(* IEC 61131-3 sources: kns-pump-station/tests/POUs/Station/FB_ControlSelector_Test, 6 files *)

(* ---- ChangedPulsesOnce.method.decl.st ---- *)
// xChanged — один вызов на смену управления (вход без рывка); без смены — FALSE
METHOD PRIVATE ChangedPulsesOnce
VAR
    fbDut : FB_ControlSelector;          // ФБ под тестом
END_VAR

(* ---- GarbageMethodIsStepped.method.decl.st ---- *)
// Способ вне перечисления — как «Ступенчатое» (E_ControlMethod: безопасный вариант)
METHOD PRIVATE GarbageMethodIsStepped
VAR
    fbDut : FB_ControlSelector;          // ФБ под тестом
    pRaw : POINTER TO INT;             // способ вне перечисления
    eBad  : E_ControlMethod;            // мусор
END_VAR

(* ---- ManualModeAlwaysManual.method.decl.st ---- *)
// 04 §4: в «Ручном» — Manual при любых условиях (защиты действуют блокировками, без запросов); режим вне
// перечисления — как «Ручной»
METHOD PRIVATE ManualModeAlwaysManual
VAR
    fbDut : FB_ControlSelector;          // ФБ под тестом
    pRaw : POINTER TO INT;             // режим вне перечисления
    eBad  : E_StationMode;              // мусор
END_VAR

(* ---- PidNotReadyFallsBackToStepped.method.decl.st ---- *)
// 04 §7.4, PMI-28: выбран ПИД, ПИД не готов — Stepped и условие KNS1.STEP; готов — LevelPid без условия
METHOD PRIVATE PidNotReadyFallsBackToStepped
VAR
    fbDut : FB_ControlSelector;          // ФБ под тестом
END_VAR

(* ---- PrecedenceTable.method.decl.st ---- *)
// 04 §4: старшинство в «Автомате» PowerLost > Restart > DryRunStop > Float > Emergency > LevelPid > Stepped — для
// каждой пары условий побеждает старшее (все 2^5 сочетаний пяти условий при выбранном и готовом ПИД)
METHOD PRIVATE PrecedenceTable
VAR
    fbDut : FB_ControlSelector;          // ФБ под тестом

    uiMask   : UINT;                    // сочетание условий: бит 0 PowerLost … бит 4 Emergency
    eExpect  : E_ControlAct;            // ожидаемое управление
    xAllOk   : BOOL := TRUE;            // все сочетания дали ожидаемое
    uiBad    : UINT;                    // первое неверное сочетание
END_VAR

(* ---- PrecedenceTable.method.impl.st ---- *)
coUnit.TEST('ControlSelector_PrecedenceTable_A4');

FOR uiMask := 0 TO 31 DO
    fbDut(eMode := E_StationMode.Auto, eMethod := E_ControlMethod.LevelPid, xPowerLost := (uiMask AND 1) <> 0,
          xRestart := (uiMask AND 2) <> 0, xDryRun := (uiMask AND 4) <> 0, xFloatMode := (uiMask AND 8) <> 0,
          xEmergency := (uiMask AND 16) <> 0, xPidReady := TRUE);
    IF (uiMask AND 1) <> 0 THEN
        eExpect := E_ControlAct.PowerLost;
    ELSIF (uiMask AND 2) <> 0 THEN
        eExpect := E_ControlAct.Restart;
    ELSIF (uiMask AND 4) <> 0 THEN
        eExpect := E_ControlAct.DryRunStop;
    ELSIF (uiMask AND 8) <> 0 THEN
        eExpect := E_ControlAct.Float;
    ELSIF (uiMask AND 16) <> 0 THEN
        eExpect := E_ControlAct.Emergency;
    ELSE
        eExpect := E_ControlAct.LevelPid;
    END_IF
    IF fbDut.eControlAct <> eExpect AND xAllOk THEN
        xAllOk := FALSE;
        uiBad := uiMask;
    END_IF
END_FOR
AssertTrue(Condition := xAllOk, Message := 'precedence: higher condition always wins');
AssertEquals_UINT(Expected := 0, Actual := uiBad, Message := 'first wrong combination');
fbDut(eMode := E_StationMode.Auto, eMethod := E_ControlMethod.Stepped, xPowerLost := FALSE, xRestart := FALSE,
      xDryRun := FALSE, xFloatMode := FALSE, xEmergency := FALSE, xPidReady := TRUE);
AssertTrue(Condition := fbDut.eControlAct = E_ControlAct.Stepped, Message := 'nothing active, Stepped selected');

coUnit.TEST_FINISHED();
